Fanuc KAREL source: kd00076.KL

-- PROVISIONAL review KL for V1013-1; original PC SHA256 481c27a82db9f692b490a3f6e1298dcde38d9a1ee1d90e673aa59a5bb66a374f
-- Incomplete behavior may be omitted. Consult companion uncertainty JSON. Do not deploy.
PROGRAM KD00076
%NOLOCKGROUP
VAR
  I : INTEGER
  J : INTEGER
  B : BOOLEAN
  R : REAL
  S : STRING[80]
BEGIN
  -- UNRESOLVED_PC offsets 5-7; opcodes 9D,3C
  -- UNRESOLVED_PC offsets 12-16; opcodes 7F
END KD00076
